FUNCTION_BLOCK Resistance (* Composite Function Block Type *)
  (* Standard: 61499-2 *)
  (* Version 0.0, 6/21/2016, Andrei, nxtControl GmbH, template *)
  PACKAGE Main;
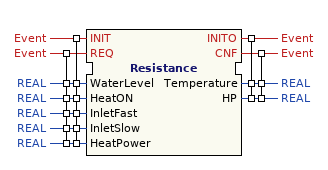
  EVENT_INPUT
    INIT WITH WaterLevel, HeatON, InletFast, InletSlow, HeatPower; (* Initialization Request *)
    REQ WITH WaterLevel, HeatON, InletFast, InletSlow, HeatPower; (* Normal Execution Request *)
  END_EVENT
  EVENT_OUTPUT
    INITO WITH Temperature, HP; (* Initialization Confirm *)
    CNF WITH Temperature, HP; (* Execution Confirmation *)
  END_EVENT
  VAR_INPUT
    WaterLevel : REAL;
    HeatON : REAL; (* Input event qualifier *)
    InletFast : REAL;
    InletSlow : REAL;
    HeatPower : REAL;
  END_VAR
  VAR_OUTPUT
    Temperature : REAL; (* Output event qualifier *)
    HP : REAL;
  END_VAR
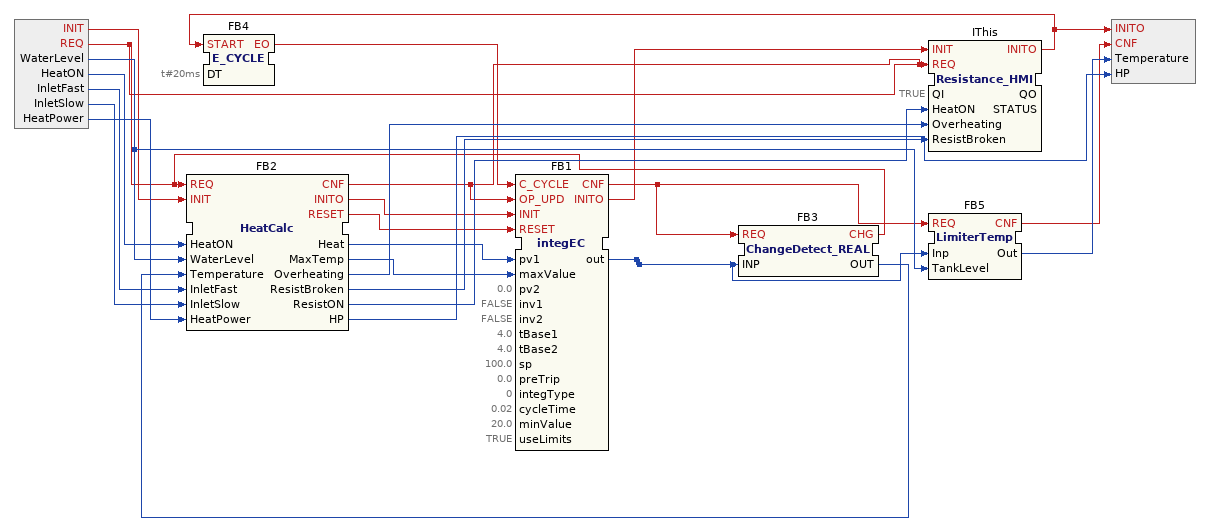
  FBS
    FB1 : integEC(pv2 := 0.0, inv1 := FALSE, inv2 := FALSE, tBase1 := 4.0, tBase2 := 4.0, sp := 100.0, preTrip := 0.0, integType := 0, cycleTime := 0.02, minValue := 20.0, useLimits := TRUE);
    FB3 : ChangeDetect_REAL;
    FB4 : E_CYCLE(DT := t#20ms);
    IThis : Resistance_HMI(QI := TRUE);
    FB5 : LimiterTemp;
    FB2 : HeatCalc;
  END_FBS
  EVENT_CONNECTIONS
    FB1.CNF TO FB3.REQ;
    FB4.EO TO FB1.C_CYCLE;
    FB2.CNF TO FB1.OP_UPD;
    FB2.INITO TO FB1.INIT;
    REQ TO FB2.REQ;
    INIT TO FB2.INIT;
    FB2.RESET TO FB1.RESET;
    FB3.CHG TO FB2.REQ;
    FB1.CNF TO FB5.REQ;
    FB5.CNF TO CNF;
    FB1.INITO TO IThis.INIT;
    REQ TO IThis.REQ;
    FB2.CNF TO IThis.REQ;
    IThis.INITO TO INITO;
    IThis.INITO TO FB4.START;
  END_CONNECTIONS
  DATA_CONNECTIONS
    HeatON TO FB2.HeatON;
    WaterLevel TO FB2.WaterLevel;
    FB2.Heat TO FB1.pv1;
    FB1.out TO FB3.INP;
    FB3.OUT TO FB2.Temperature;
    FB2.MaxTemp TO FB1.maxValue;
    FB1.out TO FB5.Inp;
    FB5.Out TO Temperature;
    FB2.Overheating TO IThis.Overheating;
    FB2.ResistBroken TO IThis.ResistBroken;
    WaterLevel TO FB5.TankLevel;
    InletFast TO FB2.InletFast;
    InletSlow TO FB2.InletSlow;
    FB2.ResistON TO IThis.HeatON;
    HeatPower TO FB2.HeatPower;
    FB2.HP TO HP;
  END_CONNECTIONS
END_FUNCTION_BLOCK
